Fanuc KAREL source: KB00001.KL

PROGRAM KB00001
%NOLOCKGROUP
%ENVIRONMENT MULTI
VAR
  P1: STRING[80]
  P2: BOOLEAN
  P3: BOOLEAN
  P4: INTEGER
BEGIN
  P1 = 'A'
  P2 = TRUE
  P3 = TRUE
  P4 = 1
  ABORT_TASK(P1, P2, P3, P4)
END KB00001
